            num nMoveType = 1
            num nPercentage
            num nSigValue = 1
        pointRx pPointRx[2] = {x=31.939332, y=-335.340311, z=740.403694, rx=-3.0192557, ry=-0.381221, rz=179.995993, shoulder=lefty, elbow=enegative, wrist=wnegative}
        string sID
      [34]
        bool bMarked
        jointRx jJointRx = {j1=-84.237822, j2=115.317662, j3=-121.0776042, j4=178.411151, j5=-2.718919, j6=85.828868}
        pointRx pInter
        paraItem pParaItem
          [0]
            bool bSafePoint
            ifItem iIfItem
              [0]
                bool bANDOR[2]
                num nSigIndex[3]
                num nSigType[3]
                num nValue[3]
            mdesc mMdesc
            num nActionIndex = 42
            num nDelay
            num nMoveType = 1
            num nPercentage
            num nSigValue = 1
        pointRx pPointRx[2] = {x=85.737999, y=-358.193052, z=740.403684, rx=-3.0191687, ry=-0.38026, rz=179.995965, shoulder=lefty, elbow=enegative, wrist=wnegative}
        string sID
      [35]
        bool bMarked
        jointRx jJointRx = {j1=-82.00566217, j2=112.688592, j3=-130.317472, j4=180.166039, j5=-14.585147, j6=81.852348}
        pointRx pInter
        paraItem pParaItem
          [0]
            bool bSafePoint
            ifItem iIfItem
              [0]
                bool bANDOR[2]
                num nSigIndex[3]
                num nSigType[3]
                num nValue[3]
            mdesc mMdesc
            num nActionIndex = 42
            num nDelay
            num nMoveType = 1
            num nPercentage
            num nSigValue = 1
        pointRx pPointRx[2] = {x=89.769203, y=-277.0582017, z=740.403696, rx=-3.0200723, ry=-0.381714, rz=179.9962, shoulder=lefty, elbow=enegative, wrist=wnegative}
        string sID
      [36]
        bool bMarked
        jointRx jJointRx = {j1=-72.862793, j2=113.115191, j3=-129.396671, j4=182.28025, j5=-13.293623, j6=70.663681}
        pointRx pInter
        paraItem pParaItem
          [0]
            bool bSafePoint
            ifItem iIfItem
              [0]
                bool bANDOR[2]
                num nSigIndex[3]
                num nSigType[3]
                num nValue[3]
            mdesc mMdesc
            num nActionIndex = 42
            num nDelay
            num nMoveType = 1
            num nPercentage
            num nSigValue = 1
        pointRx pPointRx[2] = {x=139.246931, y=-266.374782, z=740.403649, rx=-3.0193988, ry=-0.382047, rz=179.996313, shoulder=lefty, elbow=enegative, wrist=wnegative}
        string sID
      [37]
        bool bMarked
        jointRx jJointRx = {j1=-62.25584, j2=114.51749, j3=-125.317693, j4=187.673812, j5=-8.0201105, j6=54.689044}
        pointRx pInter
        paraItem pParaItem
          [0]
            bool bSafePoint
            ifItem iIfItem
              [0]
                bool bANDOR[2]
                num nSigIndex[3]
                num nSigType[3]
                num nValue[3]
            mdesc mMdesc
            num nActionIndex = 42
            num nDelay
            num nMoveType = 1
            num nPercentage
            num nSigValue = 1
        pointRx pPointRx[2] = {x=207.132214, y=-266.374817, z=740.40358, rx=-3.0201446, ry=-0.381695, rz=179.996214, shoulder=lefty, elbow=enegative, wrist=wnegative}
        string sID
      [38]
        bool bMarked
        jointRx jJointRx = {j1=-62.25584, j2=114.51749, j3=-125.317693, j4=187.673812, j5=-8.0201105, j6=54.689044}
        pointRx pInter
        paraItem pParaItem
          [0]
            bool bSafePoint
            ifItem iIfItem
              [0]
                bool bANDOR[2]
                num nSigIndex[3]
                num nSigType[3]
                num nValue[3]
            mdesc mMdesc
            num nActionIndex = 42
            num nDelay
            num nMoveType
            num nPercentage
            num nSigValue = 1
        pointRx pPointRx[2] = {x=207.132214, y=-266.374817, z=740.40358, rx=-3.0201446, ry=-0.381695, rz=179.996214, shoulder=lefty, elbow=enegative, wrist=wnegative}
        string sID
      [39]
        bool bMarked
        jointRx jJointRx = {j1=-69.425067, j2=115.601832, j3=-118.606607, j4=144.176063, j5=0.65466, j6=105.101635}
        pointRx pInter
        paraItem pParaItem
          [0]
            bool bSafePoint
            ifItem iIfItem
              [0]
                bool bANDOR[2]
                num nSigIndex[3]
                num nSigType[3]
                num nValue[3]
            mdesc mMdesc
            num nActionIndex = 42
            num nDelay
            num nMoveType
            num nPercentage
            num nSigValue = 1
        pointRx pPointRx[2] = {x=183.541944, y=-337.16529, z=739.804177, rx=-3.445036, ry=-0.883019, rz=179.816025, shoulder=lefty, elbow=enegative, wrist=wpositive}
        string sID
      [40]
        bool bMarked
        jointRx jJointRx = {j1=-72.00363568, j2=115.150585, j3=-107.679214, j4=178.830759, j5=11.0234072, j6=73.00080801}
        pointRx pInter
        paraItem pParaItem
          [0]
            bool bSafePoint
            ifItem iIfItem
              [0]
                bool bANDOR[2]
                num nSigIndex[3]
                num nSigType[3]
                num nValue[3]
            mdesc mMdesc
            num nActionIndex = 42
            num nDelay
            num nMoveType = 1
            num nPercentage
            num nSigValue = 1
        pointRx pPointRx[2] = {x=191.224277, y=-420.505468, z=739.804144, rx=-3.445497, ry=-0.883441, rz=179.816, shoulder=lefty, elbow=enegative, wrist=wpositive}
        string sID
      [41]
        bool bMarked
        jointRx jJointRx = {j1=-63.604591, j2=115.581965, j3=-112.253643, j4=173.794215, j5=6.847684, j6=69.631443}
        pointRx pInter
        paraItem pParaItem
          [0]
            bool bSafePoint
            ifItem iIfItem
              [0]
                bool bANDOR[2]
                num nSigIndex[3]
                num nSigType[3]
                num nValue[3]
            mdesc mMdesc
            num nActionIndex = 42
            num nDelay
            num nMoveType = 1
            num nPercentage
            num nSigValue = 1
        pointRx pPointRx[2] = {x=240.684957, y=-357.988391, z=739.804111, rx=-3.445463, ry=-0.88438, rz=179.815962, shoulder=lefty, elbow=enegative, wrist=wpositive}
        string sID
      [42]
        bool bMarked
        jointRx jJointRx = {j1=-53.383634, j2=115.338258, j3=-109.311316, j4=171.755597, j5=9.415846, j6=61.399656}
        pointRx pInter
        paraItem pParaItem
          [0]
            bool bSafePoint
            ifItem iIfItem
              [0]
                bool bANDOR[2]
                num nSigIndex[3]
                num nSigType[3]
                num nValue[3]
            mdesc mMdesc
            num nActionIndex = 42
            num nDelay
            num nMoveType = 1
            num nPercentage
            num nSigValue = 1
        pointRx pPointRx[2] = {x=317.964208, y=-324.389308, z=739.804138, rx=-3.445379, ry=-0.883865, rz=179.815971, shoulder=lefty, elbow=enegative, wrist=wpositive}
        string sID
      [43]
        bool bMarked
        jointRx jJointRx = {j1=-59.402506, j2=113.338107, j3=-97.632645, j4=176.975483, j5=19.145019, j6=62.132037}
        pointRx pInter
        paraItem pParaItem
          [0]
            bool bSafePoint
            ifItem iIfItem
              [0]
                bool bANDOR[2]
                num nSigIndex[3]
                num nSigType[3]
                num nValue[3]
            mdesc mMdesc
            num nActionIndex = 42
            num nDelay
            num nMoveType = 1
            num nPercentage
            num nSigValue = 1
        pointRx pPointRx[2] = {x=317.96415, y=-422.472428, z=739.804106, rx=-3.444321, ry=-0.883491, rz=179.815889, shoulder=lefty, elbow=enegative, wrist=wpositive}
        string sID
      [44]
        bool bMarked
        jointRx jJointRx = {j1=-58.0600297, j2=108.105024, j3=-79.42328, j4=177.983092, j5=32.0883294, j6=59.642392}
        pointRx pInter
        paraItem pParaItem
          [0]
            bool bSafePoint
            ifItem iIfItem
              [0]
                bool bANDOR[2]
                num nSigIndex[3]
                num nSigType[3]
                num nValue[3]
            mdesc mMdesc
            num nActionIndex = 42
            num nDelay
            num nMoveType = 1
            num nPercentage
            num nSigValue = 1
        pointRx pPointRx[2] = {x=382.78857, y=-501.837589, z=739.816752, rx=-3.444284, ry=-0.883375, rz=179.81511, shoulder=lefty, elbow=enegative, wrist=wpositive}
        string sID
      [45]
        bool bMarked
        jointRx jJointRx = {j1=-57.462056, j2=95.846947, j3=-71.551208, j4=177.618324, j5=27.69562, j6=59.445484}
        pointRx pInter
        paraItem pParaItem
          [0]
            bool bSafePoint
            ifItem iIfItem
              [0]
                bool bANDOR[2]
                num nSigIndex[3]
                num nSigType[3]
                num nValue[3]
            mdesc mMdesc
            num nActionIndex = 42
            num nDelay
            num nMoveType = 1
            num nPercentage
            num nSigValue = 1
        pointRx pPointRx[2] = {x=382.788593, y=-489.0644454, z=843.101413, rx=-3.444553, ry=-0.883416, rz=179.815149, shoulder=lefty, elbow=enegative, wrist=wpositive}
        string sID
      [46]
        bool bMarked
        jointRx jJointRx = {j1=-52.666129, j2=89.154615, j3=-75.0738664, j4=175.366505, j5=17.41012, j6=56.969519}
        pointRx pInter
        paraItem pParaItem
          [0]
            bool bSafePoint
            ifItem iIfItem
              [0]
                bool bANDOR[2]
                num nSigIndex[3]
                num nSigType[3]
                num nValue[3]
            mdesc mMdesc
            num nActionIndex = 42
            num nDelay
            num nMoveType = 1
            num nPercentage
            num nSigValue = 1
        pointRx pPointRx[2] = {x=382.788575, y=-399.492554, z=917.538047, rx=-3.444887, ry=-0.883932, rz=179.815117, shoulder=lefty, elbow=enegative, wrist=wpositive}
        string sID
      [47]
        bool bMarked
        jointRx jJointRx = {j1=-43.60719, j2=90.831848, j3=-88.576179, j4=160.320066, j5=5.597805, j6=63.0916803}
        pointRx pInter
        paraItem pParaItem
          [0]
            bool bSafePoint
            ifItem iIfItem
              [0]
                bool bANDOR[2]
                num nSigIndex[3]
                num nSigType[3]
                num nValue[3]
            mdesc mMdesc
            num nActionIndex = 42
            num nDelay
            num nMoveType = 1
            num nPercentage
            num nSigValue = 1
        pointRx pPointRx[2] = {x=382.788892, y=-272.880308, z=917.538027, rx=-3.444134, ry=-0.884317, rz=179.815078, shoulder=lefty, elbow=enegative, wrist=wpositive}
        string sID
      [48]
        bool bMarked
        jointRx jJointRx = {j1=-54.865163, j2=112.528286, j3=-89.695146, j4=177.147223, j5=26.188051, j6=57.30371}
        pointRx pInter
        paraItem pParaItem
          [0]
            bool bSafePoint
            ifItem iIfItem
              [0]
                bool bANDOR[2]
                num nSigIndex[3]
                num nSigType[3]
                num nValue[3]
            mdesc mMdesc
            num nActionIndex = 42
            num nDelay
            num nMoveType = 1
            num nPercentage
            num nSigValue = 1
        pointRx pPointRx[2] = {x=382.788429, y=-437.986191, z=727.899206, rx=-3.445194, ry=-0.883899, rz=179.815061, shoulder=lefty, elbow=enegative, wrist=wpositive}
        string sID
      [49]
        bool bMarked
        jointRx jJointRx = {j1=-87.553471, j2=145.12737, j3=-83.0900679, j4=182.117938, j5=63.691768, j6=-64.957345}
        pointRx pInter
        paraItem pParaItem
          [0]
            bool bSafePoint
            ifItem iIfItem
              [0]
                bool bANDOR[2]
                num nSigIndex[3]
                num nSigType[3]
                num nValue[3]
            mdesc mMdesc
            num nActionIndex = 42
            num nDelay
            num nMoveType = 1
            num nPercentage
            num nSigValue = 1
        pointRx pPointRx[2] = {x=61.326125, y=-652.062172, z=350.121525, rx=-1.556374, ry=-1.966704, rz=28.428639, shoulder=lefty, elbow=enegative, wrist=wpositive}
        string sID
    string sID
  [Position8_point_wash]
    num nFrameIndex
    num nMoveID
    num nToolIndex
    pointItem pPointItem[51]
      [0]
        bool bMarked
        jointRx jJointRx
        pointRx pInter
        paraItem pParaItem
          [0]
            bool bSafePoint
            ifItem iIfItem
              [0]
                bool bANDOR[2]
                num nSigIndex[3]
                num nSigType[3]
                num nValue[3]
            mdesc mMdesc
            num nActionIndex = 41
            num nDelay
            num nMoveType = 4
            num nPercentage
            num nSigValue = 1
        pointRx pPointRx[2]
        string sID
      [1]
        bool bMarked
        jointRx jJointRx
        pointRx pInter
        paraItem pParaItem
          [0]
            bool bSafePoint
            ifItem iIfItem
              [0]
                bool bANDOR[2]
                num nSigIndex[3]
                num nSigType[3]
                num nValue[3]
            mdesc mMdesc
            num nActionIndex = 42
            num nDelay
            num nMoveType = 4
            num nPercentage
            num nSigValue = 1
        pointRx pPointRx[2]
        string sID
      [2]
        bool bMarked
        jointRx jJointRx = {j1=-87.553471, j2=145.12737, j3=-83.0900679, j4=182.117938, j5=63.691768, j6=-64.957345}
        pointRx pInter
        paraItem pParaItem
          [0]
            bool bSafePoint
            ifItem iIfItem
              [0]
                bool bANDOR[2]
                num nSigIndex[3]
                num nSigType[3]
                num nValue[3]
            mdesc mMdesc
            num nActionIndex = 42
            num nDelay
            num nMoveType = 1
            num nPercentage
            num nSigValue = 1
        pointRx pPointRx[2] = {x=61.326125, y=-652.062172, z=350.121525, rx=-1.556374, ry=-1.966704, rz=28.428639, shoulder=lefty, elbow=enegative, wrist=wpositive}
        string sID
      [3]
        bool bMarked
        jointRx jJointRx = {j1=-58.11069, j2=109.524278, j3=-71.857715, j4=179.347561, j5=40.141515, j6=-122.34843}
        pointRx pInter
        paraItem pParaItem
          [0]
            bool bSafePoint
            ifItem iIfItem
              [0]
                bool bANDOR[2]
                num nSigIndex[3]
                num nSigType[3]
                num nValue[3]
            mdesc mMdesc
            num nActionIndex = 42
            num nDelay
            num nMoveType = 1
            num nPercentage
            num nSigValue = 1
        pointRx pPointRx[2] = {x=409.39132, y=-556.393527, z=693.904783, rx=-2.322296, ry=-0.948981, rz=-0.986203, shoulder=lefty, elbow=enegative, wrist=wpositive}
        string sID
      [4]
        bool bMarked
        jointRx jJointRx = {j1=-66.225547, j2=113.999088, j3=-83.778734, j4=179.876465, j5=32.728091, j6=-114.636276}
        pointRx pInter
        paraItem pParaItem
          [0]
            bool bSafePoint
            ifItem iIfItem
              [0]
                bool bANDOR[2]
                num nSigIndex[3]
                num nSigType[3]
                num nValue[3]
            mdesc mMdesc
            num nActionIndex = 42
            num nDelay
            num nMoveType = 1
            num nPercentage
            num nSigValue = 1
        pointRx pPointRx[2] = {x=300.386557, y=-556.417777, z=693.904772, rx=-2.32202, ry=-0.949536, rz=-0.986453, shoulder=lefty, elbow=enegative, wrist=wpositive}
        string sID
      [5]
        bool bMarked
        jointRx jJointRx = {j1=-76.687433, j2=116.715992, j3=-91.802088, j4=180.847193, j5=27.394171, j6=-105.0405035}
        pointRx pInter
        paraItem pParaItem
          [0]
            bool bSafePoint
            ifItem iIfItem
              [0]
                bool bANDOR[2]
                num nSigIndex[3]
                num nSigType[3]
                num nValue[3]
            mdesc mMdesc
            num nActionIndex = 42
            num nDelay
            num nMoveType = 1
            num nPercentage
            num nSigValue = 1
        pointRx pPointRx[2] = {x=180.521932, y=-560.5436, z=693.904726, rx=-2.321521, ry=-0.949691, rz=-0.986547, shoulder=lefty, elbow=enegative, wrist=wpositive}
        string sID
      [6]
        bool bMarked
        jointRx jJointRx = {j1=-85.620281, j2=117.92465, j3=-95.696322, j4=181.846877, j5=24.627005, j6=-97.0419871}
        pointRx pInter
        paraItem pParaItem
          [0]
            bool bSafePoint
            ifItem iIfItem
              [0]
                bool bANDOR[2]
                num nSigIndex[3]
                num nSigType[3]
                num nValue[3]
            mdesc mMdesc
            num nActionIndex = 42
            num nDelay
            num nMoveType = 1
            num nPercentage
            num nSigValue = 1
        pointRx pPointRx[2] = {x=86.341042, y=-560.508796, z=693.904766, rx=-2.321719, ry=-0.949521, rz=-0.986489, shoulder=lefty, elbow=enegative, wrist=wpositive}
        string sID
      [7]
        bool bMarked
        jointRx jJointRx = {j1=-101.0757166, j2=116.15458, j3=-90.0727261, j4=182.913944, j5=28.207981, j6=-82.484873}
        pointRx pInter
        paraItem pParaItem
          [0]
            bool bSafePoint
            ifItem iIfItem
              [0]
                bool bANDOR[2]
                num nSigIndex[3]
                num nSigType[3]
                num nValue[3]
            mdesc mMdesc
            num nActionIndex = 42
            num nDelay
            num nMoveType = 1
            num nPercentage
            num nSigValue = 1
        pointRx pPointRx[2] = {x=-77.997367, y=-596.182081, z=693.904723, rx=-2.320616, ry=-0.948845, rz=-0.986256, shoulder=lefty, elbow=enegative, wrist=wpositive}
        string sID
      [8]
        bool bMarked
        jointRx jJointRx = {j1=-100.388707, j2=113.501769, j3=-82.38876, j4=182.465739, j5=33.248966, j6=-82.665703}
        pointRx pInter
        paraItem pParaItem
          [0]
            bool bSafePoint
            ifItem iIfItem
              [0]
                bool bANDOR[2]
                num nSigIndex[3]
                num nSigType[3]
                num nValue[3]
            mdesc mMdesc
            num nActionIndex = 42
            num nDelay
            num nMoveType = 1
            num nPercentage
            num nSigValue = 1
        pointRx pPointRx[2] = {x=-77.997368, y=-637.319122, z=693.904719, rx=-2.320623, ry=-0.948795, rz=-0.986246, shoulder=lefty, elbow=enegative, wrist=wpositive}
        string sID
      [9]
        bool bMarked
        jointRx jJointRx = {j1=-112.569059, j2=111.105712, j3=-75.937343, j4=182.939146, j5=36.983748, j6=-70.774258}
        pointRx pInter
        paraItem pParaItem
          [0]
            bool bSafePoint
            ifItem iIfItem
              [0]
                bool bANDOR[2]
                num nSigIndex[3]
                num nSigType[3]
                num nValue[3]
            mdesc mMdesc
            num nActionIndex = 42
            num nDelay
            num nMoveType = 1
            num nPercentage
            num nSigValue = 1
        pointRx pPointRx[2] = {x=-227.428005, y=-637.284544, z=693.904751, rx=-2.321115, ry=-0.949679, rz=-0.986554, shoulder=lefty, elbow=enegative, wrist=wpositive}
        string sID
      [10]
        bool bMarked
        jointRx jJointRx = {j1=-113.957376, j2=114.00103433, j3=-83.784205, j4=183.416468, j5=32.000017554, j6=-69.935449}
        pointRx pInter
        paraItem pParaItem
          [0]
            bool bSafePoint
            ifItem iIfItem
              [0]
                bool bANDOR[2]
                num nSigIndex[3]
                num nSigType[3]
                num nValue[3]
            mdesc mMdesc
            num nActionIndex = 42
            num nDelay
            num nMoveType = 1
            num nPercentage
            num nSigValue = 1
        pointRx pPointRx[2] = {x=-227.392618, y=-596.00613787, z=693.904773, rx=-2.322353, ry=-0.948517, rz=-0.986316, shoulder=lefty, elbow=enegative, wrist=wpositive}
        string sID
      [11]
        bool bMarked
        jointRx jJointRx = {j1=-131.107782, j2=122.205733, j3=-114.25278, j4=193.937243, j5=9.352415, j6=-63.640524}
        pointRx pInter
        paraItem pParaItem
          [0]
            bool bSafePoint
            ifItem iIfItem
              [0]
                bool bANDOR[2]
                num nSigIndex[3]
                num nSigType[3]
                num nValue[3]
            mdesc mMdesc
            num nActionIndex = 42
            num nDelay
            num nMoveType = 1
            num nPercentage
            num nSigValue = 1
        pointRx pPointRx[2] = {x=-278.571769, y=-365.527339, z=693.923849, rx=-2.325235, ry=-0.948268, rz=-0.986383, shoulder=lefty, elbow=enegative, wrist=wpositive}
        string sID
      [12]
        bool bMarked
        jointRx jJointRx = {j1=-135.395911, j2=104.707172, j3=-76.504799, j4=184.753699, j5=29.243911, j6=-49.740588}
        pointRx pInter
        paraItem pParaItem
          [0]
            bool bSafePoint
            ifItem iIfItem
              [0]
                bool bANDOR[2]
                num nSigIndex[3]
                num nSigType[3]
                num nValue[3]
            mdesc mMdesc
            num nActionIndex = 42
            num nDelay
            num nMoveType = 1
            num nPercentage
            num nSigValue = 1
        pointRx pPointRx[2] = {x=-444.435288, y=-480.130514, z=766.167371, rx=-2.324241, ry=-0.947818, rz=-0.986236, shoulder=lefty, elbow=enegative, wrist=wpositive}
        string sID
      [13]
        bool bMarked
        jointRx jJointRx = {j1=-134.796217, j2=92.950158, j3=-65.644872, j4=184.86577, j5=28.374058, j6=-50.474125}
        pointRx pInter
        paraItem pParaItem
          [0]
            bool bSafePoint
            ifItem iIfItem
              [0]
                bool bANDOR[2]
                num nSigIndex[3]
                num nSigType[3]
                num nValue[3]
            mdesc mMdesc
            num nActionIndex = 42
            num nDelay
            num nMoveType = 1
            num nPercentage
            num nSigValue = 1
        pointRx pPointRx[2] = {x=-444.435359, y=-489.966612, z=855.290958, rx=-2.324744, ry=-0.947384, rz=-0.986218, shoulder=lefty, elbow=enegative, wrist=wpositive}
        string sID
      [14]
        bool bMarked
        jointRx jJointRx = {j1=-136.173853, j2=87.871737, j3=-63.130701, j4=185.374273, j5=25.767564, j6=-49.65473}
        pointRx pInter
        paraItem pParaItem
          [0]
            bool bSafePoint
            ifItem iIfItem
              [0]
                bool bANDOR[2]
                num nSigIndex[3]
                num nSigType[3]
                num nValue[3]
            mdesc mMdesc
            num nActionIndex = 42
            num nDelay
            num nMoveType = 1
            num nPercentage
            num nSigValue = 1
        pointRx pPointRx[2] = {x=-444.435358, y=-467.674325, z=901.291627, rx=-2.325949, ry=-0.946701, rz=-0.986341, shoulder=lefty, elbow=enegative, wrist=wpositive}
        string sID
      [15]
        bool bMarked
        jointRx jJointRx = {j1=-141.164951, j2=86.59666, j3=-69.357957, j4=187.756915, j5=18.114888, j6=-47.194082}
        pointRx pInter
        paraItem pParaItem
          [0]
            bool bSafePoint
            ifItem iIfItem
              [0]
                bool bANDOR[2]
                num nSigIndex[3]
                num nSigType[3]
                num nValue[3]
            mdesc mMdesc
            num nActionIndex = 42
            num nDelay
            num nMoveType = 1
            num nPercentage
            num nSigValue = 1
        pointRx pPointRx[2] = {x=-444.435342, y=-395.0345733, z=930.658223, rx=-2.325698, ry=-0.946616, rz=-0.986323, shoulder=lefty, elbow=enegative, wrist=wpositive}
        string sID
      [16]
        bool bMarked
        jointRx jJointRx = {j1=-150.996048, j2=88.749744, j3=-81.786263, j4=199.00922873, j5=7.675391, j6=-48.828489}
        pointRx pInter
        paraItem pParaItem
          [0]
            bool bSafePoint
            ifItem iIfItem
              [0]
                bool bANDOR[2]
                num nSigIndex[3]
                num nSigType[3]
                num nValue[3]
            mdesc mMdesc
            num nActionIndex = 42
            num nDelay
            num nMoveType = 1
            num nPercentage
            num nSigValue = 1
        pointRx pPointRx[2] = {x=-444.435068, y=-278.693508, z=930.65815, rx=-2.325239, ry=-0.948289, rz=-0.986304, shoulder=lefty, elbow=enegative, wrist=wpositive}
        string sID
      [17]
        bool bMarked
        jointRx jJointRx = {j1=-136.944318, j2=108.102124, j3=-81.594441, j4=185.0858237, j5=27.496189, j6=-48.554881}
        pointRx pInter
        paraItem pParaItem
          [0]
            bool bSafePoint
            ifItem iIfItem
              [0]
                bool bANDOR[2]
                num nSigIndex[3]
                num nSigType[3]
                num nValue[3]
            mdesc mMdesc
            num nActionIndex = 42
            num nDelay
            num nMoveType = 1
            num nPercentage
            num nSigValue = 1
        pointRx pPointRx[2] = {x=-444.435337, y=-455.673073, z=747.789181, rx=-2.325621, ry=-0.946829, rz=-0.986212, shoulder=lefty, elbow=enegative, wrist=wpositive}
        string sID
      [18]
        bool bMarked
        jointRx jJointRx = {j1=-133.102266, j2=114.394979, j3=-110.124586, j4=185.156231, j5=6.735085, j6=-104.330607}
        pointRx pInter
        paraItem pParaItem
          [0]
            bool bSafePoint
            ifItem iIfItem
              [0]
                bool bANDOR[2]
                num nSigIndex[3]
                num nSigType[3]
                num nValue[3]
            mdesc mMdesc
            num nActionIndex = 42
            num nDelay
            num nMoveType = 1
            num nPercentage
            num nSigValue = 1
        pointRx pPointRx[2] = {x=-273.0764108, y=-357.254112, z=747.804416, rx=-2.192889, ry=1.224247, rz=-52.275755, shoulder=lefty, elbow=enegative, wrist=wpositive}
        string sID
      [19]
        bool bMarked
        jointRx jJointRx = {j1=-117.270513, j2=113.78497, j3=-104.717978, j4=179.481532, j5=11.577034, j6=-114.962229}
        pointRx pInter
        paraItem pParaItem
          [0]
            bool bSafePoint
            ifItem iIfItem
              [0]
                bool bANDOR[2]
                num nSigIndex[3]
                num nSigType[3]
                num nValue[3]
            mdesc mMdesc
            num nActionIndex = 42
            num nDelay
            num nMoveType = 1
            num nPercentage
            num nSigValue = 1
        pointRx pPointRx[2] = {x=-176.508441, y=-453.51729, z=747.804419, rx=-2.183299, ry=1.242081, rz=-52.719273, shoulder=lefty, elbow=enegative, wrist=wpositive}
        string sID
      [20]
        bool bMarked
        jointRx jJointRx = {j1=-109.137554, j2=109.619736, j3=-86.542307, j4=178.941557, j5=25.551631, j6=-122.640865}
        pointRx pInter
        paraItem pParaItem
          [0]
            bool bSafePoint
            ifItem iIfItem
              [0]
                bool bANDOR[2]
                num nSigIndex[3]
                num nSigType[3]
                num nValue[3]
            mdesc mMdesc
            num nActionIndex = 42
            num nDelay
            num nMoveType = 1
            num nPercentage
            num nSigValue = 1
        pointRx pPointRx[2] = {x=-144.182021, y=-580.158289, z=747.804426, rx=-2.184454, ry=1.240986, rz=-52.719545, shoulder=lefty, elbow=enegative, wrist=wpositive}
        string sID
      [21]
        bool bMarked
        jointRx jJointRx = {j1=-105.96936, j2=113.946894, j3=-105.873919, j4=176.762051, j5=10.531462, j6=-123.577788}
        pointRx pInter
        paraItem pParaItem
          [0]
            bool bSafePoint
            ifItem iIfItem
              [0]
                bool bANDOR[2]
                num nSigIndex[3]
                num nSigType[3]
                num nValue[3]
            mdesc mMdesc
            num nActionIndex = 42
            num nDelay
            num nMoveType = 1
            num nPercentage
            num nSigValue = 1
        pointRx pPointRx[2] = {x=-78.145175, y=-473.574291, z=747.804414, rx=-2.185277, ry=1.240398, rz=-52.719616, shoulder=lefty, elbow=enegative, wrist=wpositive}
        string sID
      [22]
        bool bMarked
        jointRx jJointRx = {j1=-100.135452, j2=114.341428, j3=-109.460145, j4=173.401757, j5=7.298155, j6=-126.0452472}
        pointRx pInter
        paraItem pParaItem
          [0]
            bool bSafePoint
            ifItem iIfItem
              [0]
                bool bANDOR[2]
                num nSigIndex[3]
                num nSigType[3]
                num nValue[3]
            mdesc mMdesc
            num nActionIndex = 42
            num nDelay
            num nMoveType = 1
            num nPercentage
            num nSigValue = 1
        pointRx pPointRx[2] = {x=-23.263146, y=-455.736187, z=747.804388, rx=-2.18503, ry=1.240118, rz=-52.719596, shoulder=lefty, elbow=enegative, wrist=wpositive}
        string sID
      [23]
        bool bMarked
        jointRx jJointRx = {j1=-100.135452, j2=114.341428, j3=-109.460145, j4=173.401757, j5=7.298155, j6=-126.0452472}
        pointRx pInter
        paraItem pParaItem
          [0]
            bool bSafePoint
            ifItem iIfItem
              [0]
                bool bANDOR[2]
                num nSigIndex[3]
                num nSigType[3]
                num nValue[3]
            mdesc mMdesc
            num nActionIndex = 42
            num nDelay
            num nMoveType
            num nPercentage
            num nSigValue = 1
        pointRx pPointRx[2] = {x=-23.263146, y=-455.736187, z=747.804388, rx=-2.18503, ry=1.240118, rz=-52.719596, shoulder=lefty, elbow=enegative, wrist=wpositive}
        string sID
      [24]
        bool bMarked
        jointRx jJointRx = {j1=-106.631553, j2=109.786963, j3=-134.970625, j4=184.819916, j5=-24.691551, j6=-80.199638}
        pointRx pInter
        paraItem pParaItem
          [0]
            bool bSafePoint
            ifItem iIfItem
              [0]
                bool bANDOR[2]
                num nSigIndex[3]
                num nSigType[3]
                num nValue[3]
            mdesc mMdesc
            num nActionIndex = 42
            num nDelay
            num nMoveType
            num nPercentage
            num nSigValue = 1
        pointRx pPointRx[2] = {x=-10.865105, y=-272.383063, z=740.397718, rx=0.0307126, ry=2.090166, rz=-2.46071, shoulder=lefty, elbow=enegative, wrist=wnegative}
        string sID
      [25]
        bool bMarked
        jointRx jJointRx = {j1=-81.325877, j2=110.844378, j3=-133.586221, j4=185.246198, j5=-23.174992, j6=-105.96506}
        pointRx pInter
        paraItem pParaItem
          [0]
            bool bSafePoint
            ifItem iIfItem
              [0]
                bool bANDOR[2]
                num nSigIndex[3]
                num nSigType[3]
                num nValue[3]
            mdesc mMdesc
            num nActionIndex = 42
            num nDelay
            num nMoveType = 1
            num nPercentage
            num nSigValue = 1
        pointRx pPointRx[2] = {x=110.33304, y=-272.382932, z=740.397731, rx=0.0311611, ry=2.0907781, rz=-2.460321, shoulder=lefty, elbow=enegative, wrist=wnegative}
        string sID
      [26]
        bool bMarked
        jointRx jJointRx = {j1=-96.0712223, j2=114.244351, j3=-126.542039, j4=186.250879, j5=-10.611959, j6=-41.0712755}
        pointRx pInter
        paraItem pParaItem
          [0]
            bool bSafePoint
            ifItem iIfItem
              [0]
                bool bANDOR[2]
                num nSigIndex[3]
                num nSigType[3]
                num nValue[3]
            mdesc mMdesc
            num nActionIndex = 42
            num nDelay
            num nMoveType = 1
            num nPercentage
            num nSigValue = 1
        pointRx pPointRx[2] = {x=24.601437, y=-336.239263, z=740.397725, rx=-1.61612, ry=1.32728, rz=49.00349569, shoulder=lefty, elbow=enegative, wrist=wnegative}
        string sID
      [27]
        bool bMarked
        jointRx jJointRx = {j1=-95.690534, j2=114.696488, j3=-124.883411, j4=183.926416, j5=-8.191559, j6=-21.0119831}
        pointRx pInter
        paraItem pParaItem
          [0]
            bool bSafePoint
            ifItem iIfItem
              [0]
                bool bANDOR[2]
                num nSigIndex[3]
                num nSigType[3]
                num nValue[3]
            mdesc mMdesc
            num nActionIndex = 42
            num nDelay
            num nMoveType = 1
            num nPercentage
            num nSigValue = 1
        pointRx pPointRx[2] = {x=20.559143, y=-347.136674, z=740.39771, rx=-1.949012, ry=0.755958, rz=67.186994, shoulder=lefty, elbow=enegative, wrist=wnegative}
        string sID
      [28]
        bool bMarked
        jointRx jJointRx = {j1=-100.882638, j2=115.524729, j3=-119.715858, j4=189.99726, j5=-2.166253, j6=-21.927142}
        pointRx pInter
        paraItem pParaItem
          [0]
            bool bSafePoint
            ifItem iIfItem
              [0]
                bool bANDOR[2]
                num nSigIndex[3]
                num nSigType[3]
                num nValue[3]
            mdesc mMdesc
            num nActionIndex = 42
            num nDelay
            num nMoveType = 1
            num nPercentage
            num nSigValue = 1
        pointRx pPointRx[2] = {x=-20.271174, y=-387.650591, z=740.397525, rx=-1.949817, ry=0.75764, rz=67.18662, shoulder=lefty, elbow=enegative, wrist=wnegative}
        string sID
      [29]
        bool bMarked
        jointRx jJointRx = {j1=-98.590862, j2=115.394944, j3=-120.62517, j4=152.249394, j5=-3.377524, j6=83.0398225}
        pointRx pInter
        paraItem pParaItem
          [0]
            bool bSafePoint
            ifItem iIfItem
              [0]
                bool bANDOR[2]
